(* IEC 61131-3 sources: JingjiangArm/moonboxpro_arm_8.4/Application/Application/任务列表/Main_Task/IO配置表_1/KESAI, 7 files *)

(* ---- KS_AbsEncModule_IODeal.st ---- *)
(*@CES
Name=KS_AbsEncModule_IODeal
Type=FunctionBlock
TypeGuid=6f9dac99-8de1-4efc-8465-68ac443b7d08
Guid=9bb045c4-e8bf-4c9a-97a3-f47a040507bd
HasDeclaration=True
HasImplementation=False
*)
{DECLARATION}
FUNCTION_BLOCK KS_AbsEncModule_IODeal
VAR_INPUT
	i_xInputEn:BOOL;
	i_xOutPutEn:BOOL;
	(*这些值的处理未考虑双收双放*)
	i_pdwAbsEncSinglePos_Uw:POINTER TO DWORD;
	i_pwAbsEncMultiPos_Uw:POINTER TO WORD;
	(*收料*)
	i_pdwAbsEncSinglePos_Rw:POINTER TO DWORD;
	i_pwAbsEncMultiPos_Rw:POINTER TO WORD;
	//2025.08.20.152113+
	i_pstStAbsEncIOModule_Uw:POINTER TO StAbsEncIOModule;
	i_pstStAbsEncIOModule_Rw:POINTER TO StAbsEncIOModule;

END_VAR
VAR
	wIWTest:WORD;
	wQWTest: WORD;
	byAbsEncSts: BOOL;
END_VAR

{IMPLEMENTATION}

(* ---- KS_FB_IOMAP_AIAO.st ---- *)
(*@CES
Name=KS_FB_IOMAP_AIAO
Type=FunctionBlock
TypeGuid=6f9dac99-8de1-4efc-8465-68ac443b7d08
Guid=73306708-2bb0-4f5a-afc5-16fe3701a4d7
HasDeclaration=True
HasImplementation=False
*)
{DECLARATION}
FUNCTION_BLOCK KS_FB_IOMAP_AIAO
VAR_INPUT
	i_xEn: BOOL;(*功能块使能|*)
	i_xRdInput: BOOL;(*读io输入|*)
	i_xWrOutput: BOOL;(*写io输出|*)
	i_pstStSysParam								: POINTER TO StSysParam;
	i_pastStProgMonitoring						: POINTER TO ARRAY [1..2] OF StProgMonitoring;
END_VAR
VAR_OUTPUT
	o_xEno: BOOL;(*indicated to i_xEn|*)
	o_iErNo: INT;(*0.no err\-1.bad parameter|*)
END_VAR
VAR
	//fb_KS_FB_SetAIType: KS_FB_SetAIType;
	fbKS_FB_Analog_IO_CTL: KS_FB_Analog_IO_CTL;

	byAiFilterTms_UwRw_I					:  BYTE:= 1;(*滤波次数*)
	byAiFilterTms_UwRw_II					:  BYTE:= 1;
	byAiFilterTms_IfOf_I					:  BYTE:= 1;
	byAiFilterTms_IfOf_II					:  BYTE:= 1;
	byAiFilterTms_DiaMeasure_I				:   BYTE:= 1;
	byAiFilterTms_DiaMeasure_II				:   BYTE:= 1;
END_VAR

{IMPLEMENTATION}

(* ---- KS_FB_IOMAP_Axis.st ---- *)
(*@CES
Name=KS_FB_IOMAP_Axis
Type=FunctionBlock
TypeGuid=6f9dac99-8de1-4efc-8465-68ac443b7d08
Guid=efb5e60c-ddc2-4af2-8fa3-7122a81b8f33
HasDeclaration=True
HasImplementation=False
*)
{DECLARATION}
FUNCTION_BLOCK KS_FB_IOMAP_Axis
VAR_INPUT
	i_xEn: BOOL;(*功能块使能|*)
	i_xRdInput: BOOL;(*读io输入|*)
	i_xWrOutput: BOOL;(*写io输出|*)
	i_pastStIOMap_Axis_FE						: POINTER TO ARRAY [1..MAX_UNIT_NUM] OF StIOMap_Axis_FE;(*轴io数据区域|*)
END_VAR
VAR_OUTPUT
	o_xEno										: BOOL;(*indicated to i_xEn|*)
	o_iErNo										: INT;(*0.no err\-1.bad parameter|*)
END_VAR
VAR
	afbKS_FB_IOMap_Axis							: ARRAY [1..MAX_UNIT_NUM] OF KS_FB_MapAxisIOBasic;(*色组IO配置*)
END_VAR

{IMPLEMENTATION}

(* ---- KS_FB_IOMAP_AxisExtra.st ---- *)
(*@CES
Name=KS_FB_IOMAP_AxisExtra
Type=FunctionBlock
TypeGuid=6f9dac99-8de1-4efc-8465-68ac443b7d08
Guid=25cb3679-a8c2-486d-ba47-3ef0e5e06eed
HasDeclaration=True
HasImplementation=False
*)
{DECLARATION}
FUNCTION_BLOCK KS_FB_IOMAP_AxisExtra
VAR_INPUT
	i_xEn: BOOL;(*功能块使能|*)
	i_xRdInput: BOOL;(*读io输入|*)
	i_xWrOutput: BOOL;(*写io输出|*)
	i_pastStIOMap_Axis_Extra_FE						: POINTER TO ARRAY [1..MAX_UNIT_NUM] OF StIOMap_Axis_Extra_FE;(*轴io数据区域|*)
	i_pstStSysParam	:POINTER TO StSysParam;
END_VAR
VAR_OUTPUT
	o_xEno										: BOOL;(*indicated to i_xEn|*)
	o_iErNo										: INT;(*0.no err\-1.bad parameter|*)
END_VAR
VAR
	afbKS_FB_IOMap_AxisExtra							: ARRAY [1..MAX_UNIT_NUM] OF KS_FB_MapAxisIOExtra;(*色组IO配置*)
END_VAR

{IMPLEMENTATION}

(* ---- KS_FB_IOMAP_Main.st ---- *)
(*@CES
Name=KS_FB_IOMAP_Main
Type=FunctionBlock
TypeGuid=6f9dac99-8de1-4efc-8465-68ac443b7d08
Guid=0c668eca-7e01-4c5c-8e8c-334e0a405704
HasDeclaration=True
HasImplementation=False
*)
{DECLARATION}
FUNCTION_BLOCK KS_FB_IOMAP_Main
(*主面板IO配置分A/B系和放/收牵*)
(*正常单收单放选1和2*)
(*双收双放1和2是A系的放牵收牵，3和4是B系的放牵收牵*)
(*双收双放A放B收1和4*)
VAR_INPUT
	i_xEn: BOOL;(*功能块使能|*)
	i_xRdInput: BOOL;(*读io输入|*)
	i_xWrOutput: BOOL;(*写io输出|*)
	i_pastStIOMap_Main_FE						: POINTER TO ARRAY [1..4] OF StIOMap_Main_FE;(*轴io数据区域|*)
END_VAR
VAR_OUTPUT
	o_xEno										: BOOL;(*indicated to i_xEn|*)
	o_iErNo										: INT;(*0.no err\-1.bad parameter|*)
END_VAR
VAR
	afbKS_FB_MapIO_Main						: ARRAY [1..4] OF KS_FB_MapIO_Main;(*主面板IO配置*)
END_VAR

{IMPLEMENTATION}

(* ---- KS_FB_IOMAP_UwRw.st ---- *)
(*@CES
Name=KS_FB_IOMAP_UwRw
Type=FunctionBlock
TypeGuid=6f9dac99-8de1-4efc-8465-68ac443b7d08
Guid=eaf25297-ee60-4cfe-a7a6-0e28e870e49d
HasDeclaration=True
HasImplementation=False
*)
{DECLARATION}
 FUNCTION_BLOCK KS_FB_IOMAP_UwRw
VAR_INPUT
	i_xEn: BOOL;(*功能块使能|*)
	i_xRdInput: BOOL;(*读io输入|*)
	i_xWrOutput: BOOL;(*写io输出|*)
	i_pastStIOMap_UwRw_FE_Uw					: POINTER TO ARRAY [1..2] OF StIOMap_UwRw_FE;(*轴io数据区域|*)
	i_pastStIOMap_UwRw_FE_Rw					: POINTER TO ARRAY [1..2] OF StIOMap_UwRw_FE;(*轴io数据区域|*)
END_VAR
VAR_OUTPUT
	o_xEno										: BOOL;(*indicated to i_xEn|*)
	o_iErNo										: INT;(*0.no err\-1.bad parameter|*)
END_VAR
VAR
	afbKS_FB_MapIO_UwRw_Uw						: ARRAY [1..2] OF KS_FB_MapIO_UwRw;
	afbKS_FB_MapIO_UwRw_Rw						: ARRAY [1..2] OF KS_FB_MapIO_UwRw;
END_VAR

{IMPLEMENTATION}

(* ---- KS_FB_StepDriveIODeal.st ---- *)
(*@CES
Name=KS_FB_StepDriveIODeal
Type=FunctionBlock
TypeGuid=6f9dac99-8de1-4efc-8465-68ac443b7d08
Guid=1f71f424-bbb0-4026-8d51-b5eb48be2d01
HasDeclaration=True
HasImplementation=False
*)
{DECLARATION}
FUNCTION_BLOCK KS_FB_StepDriveIODeal
VAR_INPUT
	i_xInputEn:BOOL;
	i_xOutPutEn:BOOL;
	i_pastStDigitalMicroStepDrive :POINTER TO  ARRAY [1..MAX_UNIT_NUM] OF StDigitalMicroStepDrive;
	i_pastStStepDriveIOModule:POINTER TO ARRAY [1..MAX_UNIT_NUM] OF StStepDriveIOModule;
	i_pastStEnc0410R:POINTER TO ARRAY [1..MAX_UNIT_NUM] OF StEnc0410R;
END_VAR
VAR_OUTPUT
END_VAR
VAR
	wTest: WORD;
	afbKS_FB_StepDriveIOModule: ARRAY [1..MAX_UNIT_NUM] OF KS_FB_StepDriveIOModule;
END_VAR

{IMPLEMENTATION}
